FUNCTION_BLOCK FB_Listed

END_FUNCTION_BLOCK

(* stored: Version 1.1.0.1
   POU FB_Listed: Id {00000000-0000-0000-0000-000000000001}, SpecialFunc None *)
